FUNCTION_BLOCK A2X_LAST_8 (* MERGE 8 A2X in 1 A2X (LAST WRITER WINS je Kanal, generic FB) - UP und DOWN werden unabhaengig gemerged, welcher Socket zuletzt auf dem jeweiligen Kanal geschrieben hat, gewinnt *)
  (* Standard: 61499-2; Description: Copyright (c) 2026 Meisterschulen am Ostbahnhof This program and the accompanying materials are made available under the terms of the Eclipse Public License 2.0 which is available at https://www.eclipse.org/legal/epl-2.0/ SPDX-License-Identifier: EPL-2.0 *)
  (* Version 1.0, 2026-11-06, Franz Höpfinger, Meisterschulen am Ostbahnhof, generic FB GEN_A2X_LAST (N Sockets), Verhalten in FORTE *)
  PACKAGE adapter::events::unidirectional;
  IMPORT eclipse4diac::core::GenericClassName;
  {SET_ATTRIBUTE(eclipse4diac::core::GenericClassName, 'GEN_A2X_LAST')}
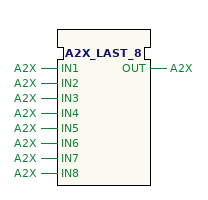
  SOCKETS
    IN1 : adapter::types::unidirectional::A2X;
    IN2 : adapter::types::unidirectional::A2X;
    IN3 : adapter::types::unidirectional::A2X;
    IN4 : adapter::types::unidirectional::A2X;
    IN5 : adapter::types::unidirectional::A2X;
    IN6 : adapter::types::unidirectional::A2X;
    IN7 : adapter::types::unidirectional::A2X;
    IN8 : adapter::types::unidirectional::A2X;
  END_SOCKETS
  PLUGS
    OUT : adapter::types::unidirectional::A2X;
  END_PLUGS
END_FUNCTION_BLOCK
